VAR_GLOBAL
	nHomingError:UDINT:=16#14D00;
END_VAR

(* stored: Version 1.1.0.1, ProductVersion 3.1.4022.6
   GVL GVL: Id {913e21aa-a47e-444c-bfce-679b16c0434b} *)
